FUNCTION_BLOCK Atuador_Coester (* Valvula com atuador Coester CSR (Modbus TCP) - HidrycoLib *)
  (* Standard: 61499-2 *)
  (* Version 2.2, 04/11/2026, Hidryco, Hidryco, 2.2: IThis.STS_ALARME (IO List da Nereda). 2.1: campo por symlink ${PATH}: mbW01..mbW09 (leitura 100 a 108), mbConexao (connStatusInt), mbCmdW01 (comando, endereco 0, em pulso) e mbCmdW02 (posicao desejada, endereco 1, so no posicionador). cfgPosicionador = TRUE: posicionar e parar (700-VC-01). Alarmes: comunicacao, falha do atuador, nao abriu/fechou/posicionou. 2.0: refeito simples. *)
  PACKAGE Hidryco.HidrycoLib;
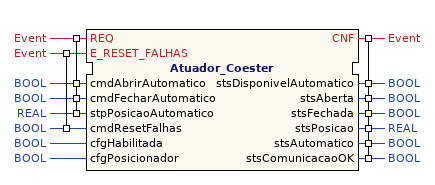
  EVENT_INPUT
    REQ WITH cmdAbrirAutomatico, cmdFecharAutomatico, stpPosicaoAutomatico; (* Atualizacao do processo *)
    E_RESET_FALHAS WITH cmdResetFalhas; (* Reset de falhas pelo processo (com cmdResetFalhas = TRUE) *)
  END_EVENT
  EVENT_OUTPUT
    CNF WITH stsDisponivelAutomatico, stsAberta, stsFechada, stsPosicao, stsAutomatico, stsComunicacaoOK; (* Status (na mudanca) *)
  END_EVENT
  VAR_INPUT
    cmdAbrirAutomatico : BOOL; (* Automatico: abrir (valvula so abrir/fechar) *)
    cmdFecharAutomatico : BOOL; (* Automatico: fechar (valvula so abrir/fechar) *)
    stpPosicaoAutomatico : REAL; (* Automatico: posicao desejada (%) - so com cfgPosicionador = TRUE *)
    cmdResetFalhas : BOOL; (* Processo: reset de falhas (vale com TRUE) *)
    cfgHabilitada : BOOL := TRUE; (* FALSE = instancia desabilitada (equipamento futuro): sem alarme de comunicacao e fora do automatico *)
    cfgPosicionador : BOOL := FALSE; (* TRUE = posicionar e parar (so 700-VC-01; o .hcf escreve tambem a Word 2, endereco 1); FALSE = so abrir e fechar *)
  END_VAR
  VAR_OUTPUT
    stsDisponivelAutomatico : BOOL; (* Pode ser comandada pelo automatico agora *)
    stsAberta : BOOL; (* Posicao aberta *)
    stsFechada : BOOL; (* Posicao fechada *)
    stsPosicao : REAL; (* Posicao real (%) - Word 5 *)
    stsAutomatico : BOOL; (* Modo automatico *)
    stsComunicacaoOK : BOOL; (* Comunicacao OK *)
  END_VAR
  FBS
    IThis : Atuador_Coester_HMI(QI := TRUE);
    plcStart1 : plcStart(Prio := 10);
    Tick : E_CYCLE(DT := T#1s);
    Leitura1 : SYMLINKMULTIVARDST_5A03F112CD5D470(QI := TRUE, NAME1 := '$${PATH}mbW01'); {SET_ATTRIBUTE(Configuration.GenericFBType.InterfaceParams, Runtime.System#I:=1;VALUE${I$}:INT)}
    Leitura2 : SYMLINKMULTIVARDST_15292F208F22048C1(QI := TRUE, NAME1 := '$${PATH}mbW02', NAME2 := '$${PATH}mbW03', NAME3 := '$${PATH}mbW04', NAME4 := '$${PATH}mbW05'); {SET_ATTRIBUTE(Configuration.GenericFBType.InterfaceParams, Runtime.System#I:=4;VALUE${I$}:INT,INT,INT,INT)}
    Leitura3 : SYMLINKMULTIVARDST_15292F208F22048C1(QI := TRUE, NAME1 := '$${PATH}mbW06', NAME2 := '$${PATH}mbW07', NAME3 := '$${PATH}mbW08', NAME4 := '$${PATH}mbW09'); {SET_ATTRIBUTE(Configuration.GenericFBType.InterfaceParams, Runtime.System#I:=4;VALUE${I$}:INT,INT,INT,INT)}
    Conexao : SYMLINKMULTIVARDST_5A03F112CD5D470(QI := TRUE, NAME1 := '$${PATH}mbConexao'); {SET_ATTRIBUTE(Configuration.GenericFBType.InterfaceParams, Runtime.System#I:=1;VALUE${I$}:INT)}
    Logica : basicValvulaCoester;
    EscritaCmd : SYMLINKMULTIVARSRC_5A03F112CD5D470(QI := TRUE, NAME1 := '$${PATH}mbCmdW01'); {SET_ATTRIBUTE(Configuration.GenericFBType.InterfaceParams, Runtime.System#I:=1;VALUE${I$}:INT)}
    EscritaPos : SYMLINKMULTIVARSRC_5A03F112CD5D470(QI := TRUE, NAME1 := '$${PATH}mbCmdW02'); {SET_ATTRIBUTE(Configuration.GenericFBType.InterfaceParams, Runtime.System#I:=1;VALUE${I$}:INT)}
    AlarmeComunicacao : ALARM_BIT(TYPE := 1, ACKTYPE_1 := 2, ACTIVE := TRUE); {SET_ATTRIBUTE(HMI.AlarmText, Atuador sem comunicação)} {SET_ATTRIBUTE(HMI.AlarmClass, Warning)}
    AlarmeAtuador : ALARM_BIT(TYPE := 1, ACKTYPE_1 := 2, ACTIVE := TRUE); {SET_ATTRIBUTE(HMI.AlarmText, Falha informada pelo atuador)}
    AlarmePosicao : ALARM_BIT(TYPE := 1, ACKTYPE_1 := 2, ACTIVE := TRUE); {SET_ATTRIBUTE(HMI.AlarmText, Válvula não chegou à posição comandada no tempo)}
  END_FBS
  EVENT_CONNECTIONS
    plcStart1.FIRST_INIT TO IThis.2EABC7344B56B5EA;
    plcStart1.REDO_INIT TO IThis.2EABC7344B56B5EA;
    IThis.E11CDC2FD3197EF0 TO Leitura1.INIT;
    Leitura1.INITO TO Leitura2.INIT;
    Leitura2.INITO TO Leitura3.INIT;
    Leitura3.INITO TO Conexao.INIT;
    Conexao.INITO TO EscritaCmd.INIT;
    EscritaCmd.INITO TO EscritaPos.INIT;
    EscritaPos.INITO TO Logica.BC3FDAAC48C266C9;
    EscritaPos.INITO TO IThis.BE814A344599F8CD;
    Logica.2C2FA7A6E9BF9047 TO Tick.START;
    Logica.2C2FA7A6E9BF9047 TO AlarmeComunicacao.INIT;
    AlarmeComunicacao.INITO TO AlarmeComunicacao.REQ_INITDATA;
    AlarmeComunicacao.CNF_INITDATA TO AlarmeComunicacao.ACTIVATE;
    AlarmeComunicacao.INITO TO AlarmeAtuador.INIT;
    AlarmeAtuador.INITO TO AlarmeAtuador.REQ_INITDATA;
    AlarmeAtuador.CNF_INITDATA TO AlarmeAtuador.ACTIVATE;
    AlarmeAtuador.INITO TO AlarmePosicao.INIT;
    AlarmePosicao.INITO TO AlarmePosicao.REQ_INITDATA;
    AlarmePosicao.CNF_INITDATA TO AlarmePosicao.ACTIVATE;
    AlarmePosicao.INITO TO plcStart1.ACK_FIRST;
    Leitura1.CNF TO Logica.907C535FA0E42403;
    Leitura2.CNF TO Logica.1122F70F08541858;
    Leitura3.CNF TO Logica.A294594AC3667AFD;
    Conexao.CNF TO Logica.45BC53B715393160;
    Tick.EO TO Logica.AEE5258FE28533BC;
    REQ TO Logica.439C5B98809C2189;
    E_RESET_FALHAS TO Logica.E0357D841C57E206;
    Logica.8A6711B6046FDA6A TO CNF;
    IThis.63B34773AE652DFD TO Logica.38061816A8BE25E9;
    IThis.71CB1D0924F3BFDA TO Logica.30AE7F49F37189A9;
    IThis.911B24FA4AD76ACA TO Logica.EC0B2AD711C1FF32;
    IThis.155C5D6A800071CB TO Logica.93A69175E8783E53;
    IThis.30C7D4C005DA551B TO Logica.3CF8A223CC6B0E4B;
    IThis.13888B810B977A05 TO Logica.0278FF007F66B823;
    IThis.F0C1E431EEC29CAD TO Logica.3A4B67BCD45EEA9F;
    IThis.F0C1E431EEC29CAD TO AlarmeComunicacao.ACK_C1;
    IThis.F0C1E431EEC29CAD TO AlarmeAtuador.ACK_C1;
    IThis.F0C1E431EEC29CAD TO AlarmePosicao.ACK_C1;
    Logica.990117E8CD2B8B73 TO IThis.481FCEE46722FF01;
    Logica.990117E8CD2B8B73 TO AlarmeComunicacao.REQ;
    Logica.990117E8CD2B8B73 TO AlarmeAtuador.REQ;
    Logica.990117E8CD2B8B73 TO AlarmePosicao.REQ;
    AlarmeComunicacao.IND_1 TO IThis.481FCEE46722FF01;
    AlarmeAtuador.IND_1 TO IThis.481FCEE46722FF01;
    AlarmePosicao.IND_1 TO IThis.481FCEE46722FF01;
    Logica.5BDBF19AA0AAE2FE TO EscritaCmd.REQ;
    Logica.5BDBF19AA0AAE2FE TO EscritaPos.REQ;
  END_CONNECTIONS
  DATA_CONNECTIONS
    Leitura1.VALUE1 TO Logica.3192419CBD3456AF;
    Leitura2.VALUE1 TO Logica.2E741C6D9D58AA99;
    Leitura2.VALUE2 TO Logica.EEA997BD3624627A;
    Leitura2.VALUE3 TO Logica.02686A07CF0DEA75;
    Leitura2.VALUE4 TO Logica.4CF28D0E5B603273;
    Leitura3.VALUE1 TO Logica.71BCBB12C2AF0796;
    Leitura3.VALUE2 TO Logica.A8A879D27B091910;
    Leitura3.VALUE3 TO Logica.5FC4C940D239F7B7;
    Leitura3.VALUE4 TO Logica.8966B61142E1C2AB;
    Conexao.VALUE1 TO Logica.93F81E7F7C459083;
    Logica.AC804A87A5A79AB2 TO EscritaCmd.VALUE1;
    Logica.4FD4131076BF837A TO EscritaPos.VALUE1;
    cmdAbrirAutomatico TO Logica.70687EF23AE88FC9;
    cmdFecharAutomatico TO Logica.F2C6EF86A9B85995;
    stpPosicaoAutomatico TO Logica.0F827E892CBAF45A;
    cmdResetFalhas TO Logica.E15FF261880BC83D;
    cfgHabilitada TO Logica.EF3C511F4EFC8BD0;
    cfgPosicionador TO Logica.CC0CBBCAA6C58448;
    Logica.99653724F6BC8F08 TO stsDisponivelAutomatico;
    Logica.E6D08F90D5C52C33 TO stsAberta;
    Logica.5DD78840DE028F7B TO stsFechada;
    Logica.B46169A18CD32F7C TO stsPosicao;
    Logica.C86F8A1F62826E46 TO stsAutomatico;
    Logica.BCCB0E0F9BF49DCB TO stsComunicacaoOK;
    IThis.53A3AB6327E89C55 TO Logica.FE01ADD91E2DE6AA;
    IThis.782E32D396726508 TO Logica.5541C75939BAAAF4;
    IThis.25AE4D0A97EEDA36 TO Logica.C1B1DDD6702777D0;
    IThis.00ADEFE9AF996DF4 TO Logica.9314A77CB5285DA8;
    IThis.D18E1EEBEE97BF05 TO Logica.7957616432A80571;
    IThis.71ABA80F1E8A7A1D TO Logica.06F0657BBA388BF2;
    IThis.8ABE92B23ED26038 TO Logica.544203CD781FBA82;
    IThis.9FC046F40A62517B TO Logica.5D2134F1C8188850;
    IThis.95CEB40D72985F2C TO Logica.6DD97D51A927EFDE;
    IThis.4BBF2344676F45C3 TO Logica.33A1A871455C269D;
    Logica.BCCB0E0F9BF49DCB TO IThis.B969FCDEF96130B5;
    Logica.08539AB6A2423C74 TO IThis.3445C45C8D3C07B1;
    Logica.C659D358952CD6B7 TO IThis.C3A21C41518F8C92;
    Logica.85BCBF8B868D0FA4 TO IThis.56BCE793160E4F9B;
    Logica.75E55D8876A4AB2E TO IThis.E869DDA43722D98D;
    Logica.E6D08F90D5C52C33 TO IThis.585941C85BCE83DA;
    Logica.5DD78840DE028F7B TO IThis.118709CAD5681177;
    Logica.32153BE2C861ECF0 TO IThis.4D2B4ABC1DF87081;
    Logica.9AABFB91073A915A TO IThis.8BD21E91EDBEE9FF;
    Logica.D71B40294CEB30AA TO IThis.DEDA62E0EBADEB17;
    Logica.C86F8A1F62826E46 TO IThis.0DA1E5C3B5E4734A;
    Logica.99653724F6BC8F08 TO IThis.683B1DD33BEC1F11;
    Logica.A7375D096F25E9A0 TO IThis.3C283C97FD003068;
    Logica.332B35E709843BAF TO IThis.EAB8CECDEE47F405;
    Logica.B46169A18CD32F7C TO IThis.E92EDC6467677974;
    Logica.3B6F475C569C5069 TO IThis.53B5F5D2A95335A0;
    Logica.1E38EF76B7197DEE TO IThis.CAA9E8865AA9CC43;
    Logica.46F7138E9A587B4E TO IThis.A6CED4D4BB171668;
    Logica.F1568A13AC3AEFBE TO IThis.F8D90F2913DF52AF;
    Logica.A99EAB43BF4ADEB5 TO IThis.2BAF0C38CF5B5251;
    Logica.EE389DE2DBE99516 TO IThis.DC69038179C46D37;
    Logica.71F9AE205389F66A TO IThis.F9AC7CF3C819F645;
    Logica.DB7EA302241EF8BC TO IThis.DA6223C9ED3732BE;
    Logica.51C9C3E1B4E288BC TO IThis.0CDC22B197562BCC;
    Logica.7A82F28321EB8D2C TO IThis.2D2E2A67F151864E;
    Logica.08539AB6A2423C74 TO AlarmeComunicacao.INP;
    Logica.1E38EF76B7197DEE TO AlarmeAtuador.INP;
    Logica.A7375D096F25E9A0 TO AlarmePosicao.INP;
    AlarmeComunicacao.STATE_1 TO IThis.B89204E4643E3E78;
    AlarmeAtuador.STATE_1 TO IThis.E687D663B06D7C72;
    AlarmePosicao.STATE_1 TO IThis.C3B11476CBB5BCEC;
    Logica.2B816C29C7AA4CF1 TO IThis.661CD66C2E0B4EB7;
  END_CONNECTIONS
END_FUNCTION_BLOCK
